// TIA Portal V21 export
// export: Created 2026-11-07T14:35:57.2666808Z, ExportSetting WithDefaults, DisplayName Totally Integrated Automation Portal, DisplayVersion V21, DisplayName STEP 7 Professional, DisplayVersion V21, DisplayName STEP 7 Safety, DisplayVersion V21, DisplayName Tech WebApplication, DisplayVersion V21, DisplayName WinCC Basic/Comfort/Advanced, DisplayVersion V21, DisplayName WinCC Unified, DisplayVersion V21
Screen "Screen_1"  1024x768, Number=1
  ScreenLayer 
    TextField "Text field_1" at 20,17 size 95x22  Text="PLC+ 2019:"
    IOField "I/O field_1" at 86,66 size 96x32  DataFormat=Decimal, FormatPattern=s999999999.999, Mode=InOutput
      ProcessValue := time
